SUBAPPLICATION logiBUS_AI_Raw_AR_OPC (* logiBUS_AI_IDA Rohwert als AR + OPC-UA-Publish (ohne VT) *)
  (* Standard: 61499-2; Description: Copyright (c) 2026 Meisterschulen am Ostbahnhof This program and the accompanying materials are made available under the terms of the Eclipse Public License 2.0 which is available at https://www.eclipse.org/legal/epl-2.0/ SPDX-License-Identifier: EPL-2.0 *)
  (* Version 1.0, 2026-10-28, Franz Höpfinger, Meisterschulen am Ostbahnhof, Kopie von MyLib::sys::logiBUS_AI_Raw_VT_AR_OPC ohne Q_NumericValue_RAW/AUDI_SPLIT_2, fuer Stationen ohne VT (keine isobus_UT-Libs). *)
  PACKAGE MyLib::sys;
  IMPORT logiBUS::io::AI::logiBUS_AI;
  IMPORT logiBUS::io::AI::logiBUS_AI_S;
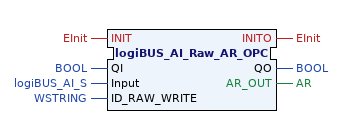
  EVENT_INPUT
    INIT : EInit; (* Initialization Request *)
  END_EVENT
  EVENT_OUTPUT
    INITO : EInit; (* Initialization Confirm *)
  END_EVENT
  VAR_INPUT
    QI : BOOL := TRUE; (* Quality Input - TRUE to enable service *)
    Input : logiBUS::io::AI::logiBUS_AI_S := logiBUS_AI::Invalid; (* Identify the Input AnalogInput_I1..I8 *)
    ID_RAW_WRITE : WSTRING; (* Rohwert-Ruckmelde-Adresse (REAL 0-4095, ACTION=PUBLISH) *)
  END_VAR
  VAR_OUTPUT
    QO : BOOL; (* Quality Output - TRUE if service executed successfully *)
  END_VAR
  PLUGS
    AR_OUT : adapter::types::unidirectional::AR; (* Rohwert als AR, fertig fuer CALIBRATE.X *)
  END_PLUGS
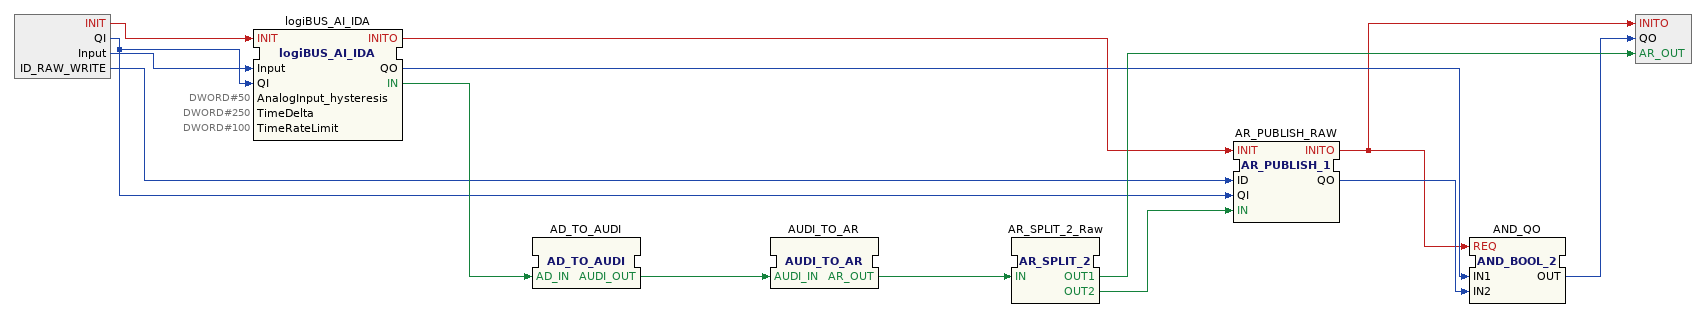
  FBS
    logiBUS_AI_IDA : logiBUS::io::AI::logiBUS_AI_IDA(AnalogInput_hysteresis := DWORD#50, TimeDelta := DWORD#250, TimeRateLimit := DWORD#100);
    AD_TO_AUDI : adapter::conversion::unidirectional::AD_TO_AUDI;
    AUDI_TO_AR : adapter::conversion::unidirectional::AUDI_TO_AR;
    AR_SPLIT_2_Raw : adapter::events::unidirectional::AR_SPLIT_2;
    AR_PUBLISH_RAW : adapter::net::AR_PUBLISH_1;
    AND_QO : iec61131::booleanOperators::AND_BOOL_2;
  END_FBS
  EVENT_CONNECTIONS
    INIT TO logiBUS_AI_IDA.INIT;
    logiBUS_AI_IDA.INITO TO AR_PUBLISH_RAW.INIT;
    AR_PUBLISH_RAW.INITO TO INITO;
    AR_PUBLISH_RAW.INITO TO AND_QO.REQ;
  END_CONNECTIONS
  DATA_CONNECTIONS
    Input TO logiBUS_AI_IDA.Input;
    ID_RAW_WRITE TO AR_PUBLISH_RAW.ID;
    QI TO logiBUS_AI_IDA.QI;
    QI TO AR_PUBLISH_RAW.QI;
    logiBUS_AI_IDA.QO TO AND_QO.IN1;
    AR_PUBLISH_RAW.QO TO AND_QO.IN2;
    AND_QO.OUT TO QO;
  END_CONNECTIONS
  ADAPTER_CONNECTIONS
    logiBUS_AI_IDA.IN TO AD_TO_AUDI.AD_IN;
    AD_TO_AUDI.AUDI_OUT TO AUDI_TO_AR.AUDI_IN;
    AUDI_TO_AR.AR_OUT TO AR_SPLIT_2_Raw.IN;
    AR_SPLIT_2_Raw.OUT1 TO AR_OUT;
    AR_SPLIT_2_Raw.OUT2 TO AR_PUBLISH_RAW.IN;
  END_CONNECTIONS
END_SUBAPPLICATION
